// TwinSAFE group diagnostic codes (EL/EJ6910).
{attribute 'qualified_only'}
{attribute 'to_string'}
TYPE
E_SafeGroupDiag :
(
    NoError := 0,
    FbError := 1,
    ComError := 2,
    ModuleError := 3,
    CmpError := 4,
    DeactivateError := 5,
    RestartError := 6
) BYTE;
END_TYPE

(* stored: Version 1.1.0.1
   DUT E_SafeGroupDiag: Id {e3bf3d65-0258-5f4b-9d53-f18cd69a8bac} *)
